(* IEC 61131-3 sources: trust-platform/examples/OSCAT/energy_normalization/non-oop/src, 3 files *)

(* ---- Configuration.st ---- *)
CONFIGURATION EnergyNormalizationClassicConfiguration
RESOURCE EnergyNormalizationClassic ON PLC
    TASK MainTask (INTERVAL := T#100ms, PRIORITY := 1);
    PROGRAM Main WITH MainTask : Main;
END_RESOURCE
END_CONFIGURATION

(* ---- Main.st ---- *)
PROGRAM Main
VAR
    EnergyConversion : ENERGY;
    SpeedConversion : SPEED;
    EnergyJoules : REAL := REAL#3600.0;
    SpeedMetersPerSecond : REAL := REAL#10.0;
    EnergyWattHours : REAL;
    SpeedKilometersPerHour : REAL;
END_VAR

EnergyConversion(J := EnergyJoules);
SpeedConversion(ms := SpeedMetersPerSecond);
EnergyWattHours := EnergyConversion.YWh;
SpeedKilometersPerHour := SpeedConversion.Ykmh;
END_PROGRAM

(* ---- Tests.st ---- *)
TEST_PROGRAM EnergyNormalizationClassicUsesConversionBlocks
VAR
    EnergyConversion : ENERGY;
    SpeedConversion : SPEED;
END_VAR

EnergyConversion(J := REAL#3600.0);
SpeedConversion(ms := REAL#10.0);

ASSERT_NEAR(EXPECTED := REAL#1.0, ACTUAL := EnergyConversion.YWh, DELTA := REAL#0.001);
ASSERT_NEAR(EXPECTED := REAL#36.0, ACTUAL := SpeedConversion.Ykmh, DELTA := REAL#0.001);
END_TEST_PROGRAM
